FUNCTION_BLOCK DrillDriver (* Composite Function Block Type *)
  (* Standard: 61499-2 *)
  (* Version 0.0, 7/2/2026, template *)
  PACKAGE Main;
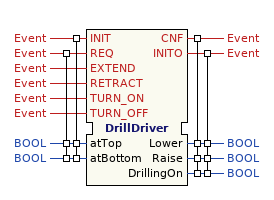
  EVENT_INPUT
    INIT WITH atTop, atBottom; (* Initialization Request *)
    REQ WITH atTop, atBottom; (* Normal Execution Request *)
    EXTEND;
    RETRACT;
    TURN_ON;
    TURN_OFF;
  END_EVENT
  EVENT_OUTPUT
    CNF WITH Lower, Raise, DrillingOn; (* Execution Confirmation *)
    INITO WITH Lower, Raise, DrillingOn; (* Initialization Confirm *)
  END_EVENT
  VAR_INPUT
    atTop : BOOL; (* Input event qualifier *)
    atBottom : BOOL;
  END_VAR
  VAR_OUTPUT
    Lower : BOOL; (* Output event qualifier *)
    Raise : BOOL;
    DrillingOn : BOOL;
  END_VAR
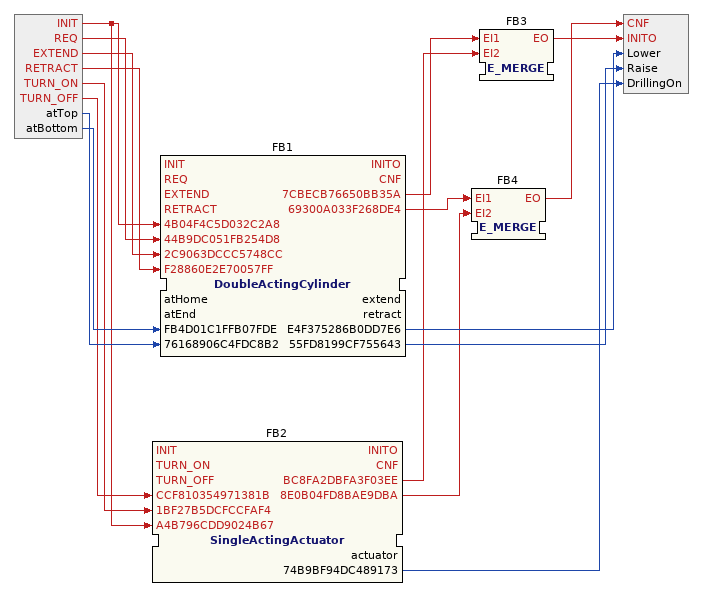
  FBS
    FB1 : DoubleActingCylinder;
    FB2 : SingleActingActuator;
    FB3 : E_MERGE;
    FB4 : E_MERGE;
  END_FBS
  EVENT_CONNECTIONS
    TURN_OFF TO FB2.CCF810354971381B;
    TURN_ON TO FB2.1BF27B5DCFCCFAF4;
    INIT TO FB2.A4B796CDD9024B67;
    INIT TO FB1.4B04F4C5D032C2A8;
    REQ TO FB1.44B9DC051FB254D8;
    EXTEND TO FB1.2C9063DCCC5748CC;
    RETRACT TO FB1.F28860E2E70057FF;
    FB4.EO TO INITO;
    FB3.EO TO CNF;
    FB1.7CBECB76650BB35A TO FB3.EI1;
    FB1.69300A033F268DE4 TO FB4.EI1;
    FB2.BC8FA2DBFA3F03EE TO FB3.EI2;
    FB2.8E0B04FD8BAE9DBA TO FB4.EI2;
  END_CONNECTIONS
  DATA_CONNECTIONS
    FB1.E4F375286B0DD7E6 TO Lower;
    FB1.55FD8199CF755643 TO Raise;
    FB2.74B9BF94DC489173 TO DrillingOn;
    atBottom TO FB1.FB4D01C1FFB07FDE;
    atTop TO FB1.76168906C4FDC8B2;
  END_CONNECTIONS
END_FUNCTION_BLOCK
